Fanuc KAREL source: KA00010.KL

PROGRAM KA00010
%NOLOCKGROUP
VAR
  SRC: INTEGER
  DST: CONFIG
BEGIN
  SRC = 2
  DST = SRC
END KA00010
